(* IEC 61131-3 sources: plc-iiot-stack/src/POUs/Iiot/F_IiotQualityText, 2 files *)

(* ---- F_IiotQualityText.decl.st ---- *)
// Назначение: текст качества для поля quality: good, uncertain, bad.
// Автор:      kr0nsch
// Версия:     0.1.0
// Документ:   docs/plc_mqtt.md, раздел «Телеметрия»
FUNCTION F_IiotQualityText : STRING(GVL_Const.IIOT_TEXT_LEN)
VAR_INPUT
    eQuality : E_IiotQuality;
END_VAR

(* ---- F_IiotQualityText.impl.st ---- *)
CASE eQuality OF
    E_IiotQuality.Good:
        F_IiotQualityText := 'good';
    E_IiotQuality.Uncertain:
        F_IiotQualityText := 'uncertain';
ELSE
    F_IiotQualityText := 'bad';
END_CASE
